// TIA Portal V20 export
// export: Created 2026-11-17T20:25:59.900199Z, ExportSetting WithDefaults, DisplayName Totally Integrated Automation Portal, DisplayVersion V20 Update 7, DisplayName TIA Portal Openness, DisplayVersion V20 Update 7, DisplayName TIA Portal Version Control Interface, DisplayVersion V20 Update 7, DisplayName TIA Portal Test Suite Advanced, DisplayVersion V20, DisplayName SINAMICS Startdrive Advanced, DisplayVersion V20 SP1 Update 1, DisplayName SINAMICS Startdrive G110M, G120, G120C, G120D, G120P, G115D, DisplayVersion V20 SP1 Update 1, DisplayName SINAMICS Startdrive G130, G150, S120, S150, SINAMICS MV, G220, S200, S210, DisplayVersion V20 SP1 Update 1, DisplayName STEP 7 Professional, DisplayVersion V20 Update 7, DisplayName STEP 7 Safety, DisplayVersion V20 Update 2, DisplayName WinCC Basic/Comfort/Advanced, DisplayVersion V20 Update 7, DisplayName WinCC Unified, DisplayVersion V20 Update 7
FUNCTION_BLOCK "zzBenTimers"   // FB240, LAD
{ S7_Optimized_Access := 'TRUE' }
VERSION : 0.1
// Benchmark networks, timers, counters, edges
// stored: AutoNumber true, IsIECCheckEnabled false, IsRetainMemResEnabled false, MemoryReserve 100, SetENOAutomatically false, UDAEnableTagReadback false
   VAR_INPUT
      inAuto : Bool;
      inLevel : Int;
      inManual : Bool;
      inSensorA : Bool;
      inSpeed : Int;
      inStart : Bool;
   END_VAR
   VAR_OUTPUT
      outQ1 : Bool;
      outQ2 : Bool;
      outQ3 : Bool;
      outQ4 : Bool;
   END_VAR
   VAR
      instCtu { S7_SetPoint := 'True'} : CTU_INT;
      instCtuA { S7_SetPoint := 'True'} : CTU_INT;
      instTonA { S7_SetPoint := 'True'} : TON_TIME;
      instTonB { S7_SetPoint := 'True'} : TON_TIME;
      statEdge : Bool;
      statElapsed : Time;
      statHold : Bool;
      statStep : Int;
   END_VAR
   VAR_TEMP   // added for the SCL form of the ladder/FBD networks
      _w1 : Bool;
   END_VAR
BEGIN

REGION Network 1: 14 Counter with fed pins
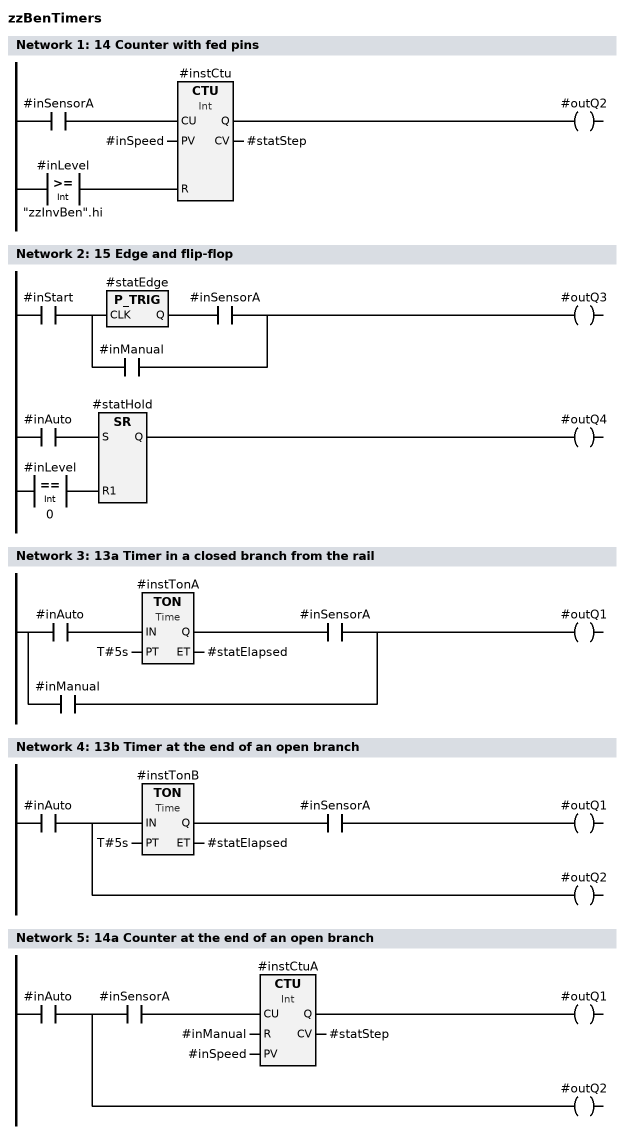
   RUNG wire#powerrail
      Contact( #inSensorA )
      { S7_Templates := "value_type := Int" } #instCtu.CTU(pv := #inSpeed, cv => #statStep, r := wire#w1)
      Coil( #outQ2 )
   END_RUNG
   RUNG wire#powerrail
      { S7_Templates := "SrcType := Int" } GE_Contact(in1 := #inLevel, in2 := "zzInvBen".hi)
   END_RUNG wire#w1
   // the same network as SCL:
   #instCtu(CU := #inSensorA, PV := #inSpeed, R := #inLevel >= "zzInvBen".hi, CV => #statStep);   // CTU
   #outQ2 := #instCtu.Q;
END_REGION

REGION Network 2: 15 Edge and flip-flop
   RUNG wire#powerrail
      Contact( #inStart )
      wire#w1
      P_Trig( #statEdge )
      Contact( #inSensorA )
      wire#w2
      Coil( #outQ3 )
   END_RUNG
   RUNG wire#w1
      Contact( #inManual )
   END_RUNG wire#w2
   RUNG wire#powerrail
      Contact( #inAuto )
      S_SR(operand := #statHold, r1 := wire#w3)
      Coil( #outQ4 )
   END_RUNG
   RUNG wire#powerrail
      { S7_Templates := "SrcType := Int" } EQ_Contact(in1 := #inLevel, in2 := 0)
   END_RUNG wire#w3
   // the same network as SCL:
   #_w1 := #inStart AND NOT #statEdge;   // rising edge
   #statEdge := #inStart;
   #outQ3 := (#_w1 AND #inSensorA) OR (#inStart AND #inManual);
   IF #inAuto THEN
       #statHold := TRUE;   // SR flip-flop
   END_IF;
   IF #inLevel = 0 THEN #statHold := FALSE; END_IF;
   #outQ4 := #statHold;
END_REGION

REGION Network 3: 13a Timer in a closed branch from the rail
   RUNG wire#powerrail
      Contact( #inAuto )
      { S7_Templates := "time_type := Time" } #instTonA.TON(pt := T#5s, et => #statElapsed)
      Contact( #inSensorA )
      wire#w1
      Coil( #outQ1 )
   END_RUNG
   RUNG wire#powerrail
      Contact( #inManual )
   END_RUNG wire#w1
   // the same network as SCL:
   #instTonA(IN := #inAuto, PT := T#5s, ET => #statElapsed);   // TON
   #outQ1 := (#instTonA.Q AND #inSensorA) OR #inManual;
END_REGION

REGION Network 4: 13b Timer at the end of an open branch
   RUNG wire#powerrail
      Contact( #inAuto )
      wire#w1
      { S7_Templates := "time_type := Time" } #instTonB.TON(pt := T#5s, et => #statElapsed)
      Contact( #inSensorA )
      Coil( #outQ1 )
   END_RUNG
   RUNG wire#w1
      Coil( #outQ2 )
   END_RUNG
   // the same network as SCL:
   #instTonB(PT := T#5s, IN := #inAuto, ET => #statElapsed);   // TON
   #outQ1 := #instTonB.Q AND #inSensorA;
   #outQ2 := #inAuto;
END_REGION

REGION Network 5: 14a Counter at the end of an open branch
   RUNG wire#powerrail
      Contact( #inAuto )
      wire#w1
      Contact( #inSensorA )
      { S7_Templates := "value_type := Int" } #instCtuA.CTU(r := #inManual, pv := #inSpeed, cv => #statStep)
      Coil( #outQ1 )
   END_RUNG
   RUNG wire#w1
      Coil( #outQ2 )
   END_RUNG
   // the same network as SCL:
   #instCtuA(CU := #inAuto AND #inSensorA, R := #inManual, PV := #inSpeed, CV => #statStep);   // CTU
   #outQ1 := #instCtuA.Q;
   #outQ2 := #inAuto;
END_REGION
END_FUNCTION_BLOCK
